(* IEC 61131-3 sources: plc-vscode/tests/st/test-ready/trust-platform/examples/OSCAT/battery_energy_storage_facade/non-oop/src, 3 files *)

(* ---- Main.st ---- *)
FUNCTION_BLOCK ClassicBessCabinet
VAR
    EnabledValue : BOOL;
    AlarmCountValue : INT;
    MqttPublishReadyValue : BOOL;
    PowerCommandValue : REAL;
    FireIsolatedValue : BOOL;
END_VAR
METHOD PUBLIC Enable
EnabledValue := TRUE;
END_METHOD
METHOD PUBLIC Update : REAL
VAR_INPUT
    StateOfChargePct : REAL;
    GridPowerCommandKw : REAL;
    FireInputHealthy : BOOL;
END_VAR
IF NOT FireInputHealthy THEN
    EnabledValue := FALSE;
    FireIsolatedValue := TRUE;
    PowerCommandValue := REAL#0.0;
    AlarmCountValue := AlarmCountValue + INT#1;
    MqttPublishReadyValue := TRUE;
ELSIF EnabledValue THEN
    FireIsolatedValue := FALSE;
    PowerCommandValue := LIMIT(REAL#-250.0, GridPowerCommandKw, REAL#250.0);
END_IF;
Update := PowerCommandValue;
END_METHOD
PUBLIC PROPERTY AlarmCount : INT
GET
    AlarmCount := AlarmCountValue;
END_GET
END_PROPERTY
PUBLIC PROPERTY FireIsolated : BOOL
GET
    FireIsolated := FireIsolatedValue;
END_GET
END_PROPERTY
END_FUNCTION_BLOCK

PROGRAM Main
VAR
    Cabinet : ClassicBessCabinet;
    Power : REAL;
END_VAR
Cabinet.Enable();
Power := Cabinet.Update(StateOfChargePct := REAL#70.0, GridPowerCommandKw := REAL#120.0, FireInputHealthy := TRUE);
END_PROGRAM

(* ---- Configuration.st ---- *)
CONFIGURATION BatteryEnergyStorageFacadeClassicConfiguration
RESOURCE Cpu0 ON PLC
    TASK MainTask (INTERVAL := T#100ms, PRIORITY := 1);
    PROGRAM Cabinet WITH MainTask : Main;
END_RESOURCE
END_CONFIGURATION

(* ---- Tests.st ---- *)
TEST_PROGRAM ClassicBessHandlesFireInline
VAR
    Cabinet : ClassicBessCabinet;
END_VAR
Cabinet.Enable();
ASSERT_NEAR(EXPECTED := REAL#0.0, ACTUAL := Cabinet.Update(StateOfChargePct := REAL#70.0, GridPowerCommandKw := REAL#120.0, FireInputHealthy := FALSE), DELTA := REAL#0.001);
ASSERT_TRUE(IN := Cabinet.FireIsolated);
ASSERT_EQUAL(EXPECTED := INT#1, ACTUAL := Cabinet.AlarmCount);
END_TEST_PROGRAM
